(* IEC 61131-3 sources: sis-interlock-demo/tests/POUs/Generated/FB_CemGen01_Test, 41 files *)

(* ---- FB_CemGen01_Test.decl.st ---- *)
// AUTO-GENERATED by cemgen 1.0.0 — не редактировать: правьте матрицу и запустите
//   python -m cemgen generate <файл матрицы .csv или .xlsx>
// Матрица: SIS-V101-CEM, объект V-101, ревизия B от 2026-10-19, SHA-256 сетки df2ed4841a9453ca
// Назначение: набор coUnit: сценарии по матрице SIS-V101-CEM, тесты 1–40 (DESIGN.md, 12.4).
//             Ожидаемые значения — эталонная модель cemgen. Стенд FB_SisHarness — по экземпляру на
//             тест.
// Автор:      kr0nsch; код — генератор cemgen
// Версия:     1.0.0
// Документ:   docs/DESIGN.md, раздел «10. Генератор cemgen»; docs/cause_effect_matrix.md
// ВНИМАНИЕ:   код демонстрационный и не предназначен для систем безопасности. Реальная ПАЗ требует
//             определения SIL, сертифицированных аппаратных и программных средств и валидации по
//             ГОСТ Р МЭК 61511.
FUNCTION_BLOCK FB_CemGen01_Test EXTENDS coUnit.FB_TestSuite
VAR
    fbH001 : FB_SisHarness;   // Matrix_PSHH101Demand_TripsOwnEffects
    fbH002 : FB_SisHarness;   // Matrix_PSHH101Delay_TripsExactlyAtDelay
    fbH003 : FB_SisHarness;   // Matrix_PSHH101Override_Denied
    fbH004 : FB_SisHarness;   // Matrix_PSHH101Reset_OnlyAfterClear
    fbH005 : FB_SisHarness;   // Matrix_PSHH101ChannelInvalid_MatchesPolicy
    fbH006 : FB_SisHarness;   // Matrix_PSHH101Bypass_ExpiresBackToVoting
    fbH007 : FB_SisHarness;   // Matrix_PSLL101Demand_TripsOwnEffects
    fbH008 : FB_SisHarness;   // Matrix_PSLL101Delay_TripsExactlyAtDelay
    fbH009 : FB_SisHarness;   // Matrix_PSLL101Override_ExpiresThenTrips
    fbH010 : FB_SisHarness;   // Matrix_PSLL101Override_ClearsAfterConfirm
    fbH011 : FB_SisHarness;   // Matrix_PSLL101Override_DemandBackRestartsConfirm
    fbH012 : FB_SisHarness;   // Matrix_PSLL101Override_ExpiryBoundsConfirm
    fbH013 : FB_SisHarness;   // Matrix_PSLL101Override_ClearedThenDelayTrips
    fbH014 : FB_SisHarness;   // Matrix_PSLL101Reset_OnlyAfterClear
    fbH015 : FB_SisHarness;   // Matrix_PSLL101ChannelInvalid_MatchesPolicy
    fbH016 : FB_SisHarness;   // Matrix_PSLL101Bypass_ExpiresBackToVoting
    fbH017 : FB_SisHarness;   // Matrix_LSHH102Demand_TripsOwnEffects
    fbH018 : FB_SisHarness;   // Matrix_LSHH102Delay_TripsExactlyAtDelay
    fbH019 : FB_SisHarness;   // Matrix_LSHH102Override_Denied
    fbH020 : FB_SisHarness;   // Matrix_LSHH102Reset_OnlyAfterClear
    fbH021 : FB_SisHarness;   // Matrix_LSHH102ChannelInvalid_MatchesPolicy
    fbH022 : FB_SisHarness;   // Matrix_LSHH102Bypass_ExpiresBackToVoting
    fbH023 : FB_SisHarness;   // Matrix_LSLL102Demand_TripsOwnEffects
    fbH024 : FB_SisHarness;   // Matrix_LSLL102Delay_TripsExactlyAtDelay
    fbH025 : FB_SisHarness;   // Matrix_LSLL102Override_ExpiresThenTrips
    fbH026 : FB_SisHarness;   // Matrix_LSLL102Override_ClearsAfterConfirm
    fbH027 : FB_SisHarness;   // Matrix_LSLL102Override_DemandBackRestartsConfirm
    fbH028 : FB_SisHarness;   // Matrix_LSLL102Override_ExpiryBoundsConfirm
    fbH029 : FB_SisHarness;   // Matrix_LSLL102Override_ClearedThenDelayTrips
    fbH030 : FB_SisHarness;   // Matrix_LSLL102Reset_OnlyAfterClear
    fbH031 : FB_SisHarness;   // Matrix_LSLL102ChannelInvalid_MatchesPolicy
    fbH032 : FB_SisHarness;   // Matrix_LSLL102Bypass_ExpiresBackToVoting
    fbH033 : FB_SisHarness;   // Matrix_TSHH103Demand_TripsOwnEffects
    fbH034 : FB_SisHarness;   // Matrix_TSHH103Delay_TripsExactlyAtDelay
    fbH035 : FB_SisHarness;   // Matrix_TSHH103Override_Denied
    fbH036 : FB_SisHarness;   // Matrix_TSHH103Reset_OnlyAfterClear
    fbH037 : FB_SisHarness;   // Matrix_TSHH103ChannelInvalid_MatchesPolicy
    fbH038 : FB_SisHarness;   // Matrix_TSHH103Bypass_ExpiresBackToVoting
    fbH039 : FB_SisHarness;   // Matrix_ASHH104Demand_TripsOwnEffects
    fbH040 : FB_SisHarness;   // Matrix_ASHH104Delay_TripsExactlyAtDelay
END_VAR

(* ---- ASHH104DelayTripsExactlyAtDelay.method.decl.st ---- *)
// AUTO-GENERATED by cemgen 1.0.0 — не редактировать: правьте матрицу и запустите
//   python -m cemgen generate <файл матрицы .csv или .xlsx>
// Матрица: SIS-V101-CEM, объект V-101, ревизия B от 2026-10-19, SHA-256 сетки df2ed4841a9453ca
// Назначение: тест Matrix_ASHH104Delay_TripsExactlyAtDelay набора FB_CemGen01_Test (сценарий по
//             матрице, DESIGN.md, 12.4).
// Автор:      kr0nsch; код — генератор cemgen
// Версия:     1.0.0
// Документ:   docs/DESIGN.md, раздел «10. Генератор cemgen»; docs/cause_effect_matrix.md
// ВНИМАНИЕ:   код демонстрационный и не предназначен для систем безопасности. Реальная ПАЗ требует
//             определения SIL, сертифицированных аппаратных и программных средств и валидации по
//             ГОСТ Р МЭК 61511.
// Причина 6 ASHH104: требование в t0; на t0 + 2 с − шаг не зафиксирована, следствия под напряжением;
// ровно на t0 + 2 с — зафиксирована, ltFirstOut = t0 + задержка.
METHOD PRIVATE ASHH104DelayTripsExactlyAtDelay
VAR
    xArmed : BOOL;    // стенд взведён: все следствия под напряжением после сброса
    ltT0   : LTIME;   // момент t0 по подменному времени стенда
END_VAR

(* ---- ASHH104DemandTripsOwnEffects.method.decl.st ---- *)
// AUTO-GENERATED by cemgen 1.0.0 — не редактировать: правьте матрицу и запустите
//   python -m cemgen generate <файл матрицы .csv или .xlsx>
// Матрица: SIS-V101-CEM, объект V-101, ревизия B от 2026-10-19, SHA-256 сетки df2ed4841a9453ca
// Назначение: тест Matrix_ASHH104Demand_TripsOwnEffects набора FB_CemGen01_Test (сценарий по
//             матрице, DESIGN.md, 12.4).
// Автор:      kr0nsch; код — генератор cemgen
// Версия:     1.0.0
// Документ:   docs/DESIGN.md, раздел «10. Генератор cemgen»; docs/cause_effect_matrix.md
// ВНИМАНИЕ:   код демонстрационный и не предназначен для систем безопасности. Реальная ПАЗ требует
//             определения SIL, сертифицированных аппаратных и программных средств и валидации по
//             ГОСТ Р МЭК 61511.
// Причина 6 ASHH104 (2oo3, задержка 2 с): требование AT104A, AT104B, AT104C = 12,80 мА (55 % НКПР;
// уставка ≥ 50 % НКПР) отключает ESDV101, ESDV102, P101A, P101B, H101, UA110; остальные следствия под
// напряжением; первопричина ASHH104.
METHOD PRIVATE ASHH104DemandTripsOwnEffects
VAR
    xArmed : BOOL;   // стенд взведён: все следствия под напряжением после сброса
END_VAR

(* ---- LSHH102BypassExpiresBackToVoting.method.decl.st ---- *)
// AUTO-GENERATED by cemgen 1.0.0 — не редактировать: правьте матрицу и запустите
//   python -m cemgen generate <файл матрицы .csv или .xlsx>
// Матрица: SIS-V101-CEM, объект V-101, ревизия B от 2026-10-19, SHA-256 сетки df2ed4841a9453ca
// Назначение: тест Matrix_LSHH102Bypass_ExpiresBackToVoting набора FB_CemGen01_Test (сценарий по
//             матрице, DESIGN.md, 12.4).
// Автор:      kr0nsch; код — генератор cemgen
// Версия:     1.0.0
// Документ:   docs/DESIGN.md, раздел «10. Генератор cemgen»; docs/cause_effect_matrix.md
// ВНИМАНИЕ:   код демонстрационный и не предназначен для систем безопасности. Реальная ПАЗ требует
//             определения SIL, сертифицированных аппаратных и программных средств и валидации по
//             ГОСТ Р МЭК 61511.
// Причина 3 LSHH102: ключ разрешения байпасов, байпас LT102A → Active; канал недостоверен → Bypassed,
// не сработало; на t0 + 8 ч − шаг — Active; ровно на t0 + 8 ч — Expired, BypassExpired, канал Invalid;
// далее — по эталонной модели.
METHOD PRIVATE LSHH102BypassExpiresBackToVoting
VAR
    xArmed : BOOL;           // стенд взведён: все следствия под напряжением после сброса
    stVs   : ST_VotingSts;   // копия состояния группы голосования
END_VAR

(* ---- LSHH102ChannelInvalidMatchesPolicy.method.decl.st ---- *)
// AUTO-GENERATED by cemgen 1.0.0 — не редактировать: правьте матрицу и запустите
//   python -m cemgen generate <файл матрицы .csv или .xlsx>
// Матрица: SIS-V101-CEM, объект V-101, ревизия B от 2026-10-19, SHA-256 сетки df2ed4841a9453ca
// Назначение: тест Matrix_LSHH102ChannelInvalid_MatchesPolicy набора FB_CemGen01_Test (сценарий по
//             матрице, DESIGN.md, 12.4).
// Автор:      kr0nsch; код — генератор cemgen
// Версия:     1.0.0
// Документ:   docs/DESIGN.md, раздел «10. Генератор cemgen»; docs/cause_effect_matrix.md
// ВНИМАНИЕ:   код демонстрационный и не предназначен для систем безопасности. Реальная ПАЗ требует
//             определения SIL, сертифицированных аппаратных и программных средств и валидации по
//             ГОСТ Р МЭК 61511.
// Причина 3 LSHH102 (2oo3, DegradeAvailable): канал LT102A недостоверен → действующая схема и
// срабатывание по политике деградации; если не сработало — требование на LT102B → по эталонной модели.
METHOD PRIVATE LSHH102ChannelInvalidMatchesPolicy
VAR
    xArmed : BOOL;           // стенд взведён: все следствия под напряжением после сброса
    stVs   : ST_VotingSts;   // копия состояния группы голосования
END_VAR

(* ---- LSHH102DelayTripsExactlyAtDelay.method.decl.st ---- *)
// AUTO-GENERATED by cemgen 1.0.0 — не редактировать: правьте матрицу и запустите
//   python -m cemgen generate <файл матрицы .csv или .xlsx>
// Матрица: SIS-V101-CEM, объект V-101, ревизия B от 2026-10-19, SHA-256 сетки df2ed4841a9453ca
// Назначение: тест Matrix_LSHH102Delay_TripsExactlyAtDelay набора FB_CemGen01_Test (сценарий по
//             матрице, DESIGN.md, 12.4).
// Автор:      kr0nsch; код — генератор cemgen
// Версия:     1.0.0
// Документ:   docs/DESIGN.md, раздел «10. Генератор cemgen»; docs/cause_effect_matrix.md
// ВНИМАНИЕ:   код демонстрационный и не предназначен для систем безопасности. Реальная ПАЗ требует
//             определения SIL, сертифицированных аппаратных и программных средств и валидации по
//             ГОСТ Р МЭК 61511.
// Причина 3 LSHH102: требование в t0; на t0 + 3 с − шаг не зафиксирована, следствия под напряжением;
// ровно на t0 + 3 с — зафиксирована, ltFirstOut = t0 + задержка.
METHOD PRIVATE LSHH102DelayTripsExactlyAtDelay
VAR
    xArmed : BOOL;    // стенд взведён: все следствия под напряжением после сброса
    ltT0   : LTIME;   // момент t0 по подменному времени стенда
END_VAR

(* ---- LSHH102DemandTripsOwnEffects.method.decl.st ---- *)
// AUTO-GENERATED by cemgen 1.0.0 — не редактировать: правьте матрицу и запустите
//   python -m cemgen generate <файл матрицы .csv или .xlsx>
// Матрица: SIS-V101-CEM, объект V-101, ревизия B от 2026-10-19, SHA-256 сетки df2ed4841a9453ca
// Назначение: тест Matrix_LSHH102Demand_TripsOwnEffects набора FB_CemGen01_Test (сценарий по
//             матрице, DESIGN.md, 12.4).
// Автор:      kr0nsch; код — генератор cemgen
// Версия:     1.0.0
// Документ:   docs/DESIGN.md, раздел «10. Генератор cemgen»; docs/cause_effect_matrix.md
// ВНИМАНИЕ:   код демонстрационный и не предназначен для систем безопасности. Реальная ПАЗ требует
//             определения SIL, сертифицированных аппаратных и программных средств и валидации по
//             ГОСТ Р МЭК 61511.
// Причина 3 LSHH102 (2oo3, задержка 3 с): требование LT102A, LT102B, LT102C = 16,16 мА (1,824 м;
// уставка ≥ 1,8 м) отключает ESDV101, H101, UA110; остальные следствия под напряжением; первопричина
// LSHH102.
METHOD PRIVATE LSHH102DemandTripsOwnEffects
VAR
    xArmed : BOOL;   // стенд взведён: все следствия под напряжением после сброса
END_VAR

(* ---- LSHH102OverrideDenied.method.decl.st ---- *)
// AUTO-GENERATED by cemgen 1.0.0 — не редактировать: правьте матрицу и запустите
//   python -m cemgen generate <файл матрицы .csv или .xlsx>
// Матрица: SIS-V101-CEM, объект V-101, ревизия B от 2026-10-19, SHA-256 сетки df2ed4841a9453ca
// Назначение: тест Matrix_LSHH102Override_Denied набора FB_CemGen01_Test (сценарий по матрице,
//             DESIGN.md, 12.4).
// Автор:      kr0nsch; код — генератор cemgen
// Версия:     1.0.0
// Документ:   docs/DESIGN.md, раздел «10. Генератор cemgen»; docs/cause_effect_matrix.md
// ВНИМАНИЕ:   код демонстрационный и не предназначен для систем безопасности. Реальная ПАЗ требует
//             определения SIL, сертифицированных аппаратных и программных средств и валидации по
//             ГОСТ Р МЭК 61511.
// Причина 3 LSHH102 без разрешённого обхода: ключ разрешения обходов, запрос → последнее событие
// OverrideDenied, обхода нет; требование → срабатывание после задержки.
METHOD PRIVATE LSHH102OverrideDenied
VAR
    xArmed : BOOL;          // стенд взведён: все следствия под напряжением после сброса
    stEv   : ST_SisEvent;   // последнее событие журнала
END_VAR

(* ---- LSHH102ResetOnlyAfterClear.method.decl.st ---- *)
// AUTO-GENERATED by cemgen 1.0.0 — не редактировать: правьте матрицу и запустите
//   python -m cemgen generate <файл матрицы .csv или .xlsx>
// Матрица: SIS-V101-CEM, объект V-101, ревизия B от 2026-10-19, SHA-256 сетки df2ed4841a9453ca
// Назначение: тест Matrix_LSHH102Reset_OnlyAfterClear набора FB_CemGen01_Test (сценарий по матрице,
//             DESIGN.md, 12.4).
// Автор:      kr0nsch; код — генератор cemgen
// Версия:     1.0.0
// Документ:   docs/DESIGN.md, раздел «10. Генератор cemgen»; docs/cause_effect_matrix.md
// ВНИМАНИЕ:   код демонстрационный и не предназначен для систем безопасности. Реальная ПАЗ требует
//             определения SIL, сертифицированных аппаратных и программных средств и валидации по
//             ГОСТ Р МЭК 61511.
// Причина 3 LSHH102: срабатывание; сброс при требовании → ResetDenied, блокирует LSHH102, следствия
// обесточены; норма → следствия всё ещё обесточены (фиксация); сброс → все следствия под напряжением.
METHOD PRIVATE LSHH102ResetOnlyAfterClear
VAR
    xArmed : BOOL;          // стенд взведён: все следствия под напряжением после сброса
    stEv   : ST_SisEvent;   // последнее событие журнала
END_VAR

(* ---- LSLL102BypassExpiresBackToVoting.method.decl.st ---- *)
// AUTO-GENERATED by cemgen 1.0.0 — не редактировать: правьте матрицу и запустите
//   python -m cemgen generate <файл матрицы .csv или .xlsx>
// Матрица: SIS-V101-CEM, объект V-101, ревизия B от 2026-10-19, SHA-256 сетки df2ed4841a9453ca
// Назначение: тест Matrix_LSLL102Bypass_ExpiresBackToVoting набора FB_CemGen01_Test (сценарий по
//             матрице, DESIGN.md, 12.4).
// Автор:      kr0nsch; код — генератор cemgen
// Версия:     1.0.0
// Документ:   docs/DESIGN.md, раздел «10. Генератор cemgen»; docs/cause_effect_matrix.md
// ВНИМАНИЕ:   код демонстрационный и не предназначен для систем безопасности. Реальная ПАЗ требует
//             определения SIL, сертифицированных аппаратных и программных средств и валидации по
//             ГОСТ Р МЭК 61511.
// Причина 4 LSLL102: ключ разрешения байпасов, байпас LT102A → Active; канал недостоверен → Bypassed,
// не сработало; на t0 + 8 ч − шаг — Active; ровно на t0 + 8 ч — Expired, BypassExpired, канал Invalid;
// далее — по эталонной модели.
METHOD PRIVATE LSLL102BypassExpiresBackToVoting
VAR
    xArmed : BOOL;           // стенд взведён: все следствия под напряжением после сброса
    stVs   : ST_VotingSts;   // копия состояния группы голосования
END_VAR

(* ---- LSLL102ChannelInvalidMatchesPolicy.method.decl.st ---- *)
// AUTO-GENERATED by cemgen 1.0.0 — не редактировать: правьте матрицу и запустите
//   python -m cemgen generate <файл матрицы .csv или .xlsx>
// Матрица: SIS-V101-CEM, объект V-101, ревизия B от 2026-10-19, SHA-256 сетки df2ed4841a9453ca
// Назначение: тест Matrix_LSLL102ChannelInvalid_MatchesPolicy набора FB_CemGen01_Test (сценарий по
//             матрице, DESIGN.md, 12.4).
// Автор:      kr0nsch; код — генератор cemgen
// Версия:     1.0.0
// Документ:   docs/DESIGN.md, раздел «10. Генератор cemgen»; docs/cause_effect_matrix.md
// ВНИМАНИЕ:   код демонстрационный и не предназначен для систем безопасности. Реальная ПАЗ требует
//             определения SIL, сертифицированных аппаратных и программных средств и валидации по
//             ГОСТ Р МЭК 61511.
// Причина 4 LSLL102 (2oo3, DegradeAvailable): канал LT102A недостоверен → действующая схема и
// срабатывание по политике деградации; если не сработало — требование на LT102B → по эталонной модели.
METHOD PRIVATE LSLL102ChannelInvalidMatchesPolicy
VAR
    xArmed : BOOL;           // стенд взведён: все следствия под напряжением после сброса
    stVs   : ST_VotingSts;   // копия состояния группы голосования
END_VAR

(* ---- LSLL102DelayTripsExactlyAtDelay.method.decl.st ---- *)
// AUTO-GENERATED by cemgen 1.0.0 — не редактировать: правьте матрицу и запустите
//   python -m cemgen generate <файл матрицы .csv или .xlsx>
// Матрица: SIS-V101-CEM, объект V-101, ревизия B от 2026-10-19, SHA-256 сетки df2ed4841a9453ca
// Назначение: тест Matrix_LSLL102Delay_TripsExactlyAtDelay набора FB_CemGen01_Test (сценарий по
//             матрице, DESIGN.md, 12.4).
// Автор:      kr0nsch; код — генератор cemgen
// Версия:     1.0.0
// Документ:   docs/DESIGN.md, раздел «10. Генератор cemgen»; docs/cause_effect_matrix.md
// ВНИМАНИЕ:   код демонстрационный и не предназначен для систем безопасности. Реальная ПАЗ требует
//             определения SIL, сертифицированных аппаратных и программных средств и валидации по
//             ГОСТ Р МЭК 61511.
// Причина 4 LSLL102: требование в t0; на t0 + 5 с − шаг не зафиксирована, следствия под напряжением;
// ровно на t0 + 5 с — зафиксирована, ltFirstOut = t0 + задержка.
METHOD PRIVATE LSLL102DelayTripsExactlyAtDelay
VAR
    xArmed : BOOL;    // стенд взведён: все следствия под напряжением после сброса
    ltT0   : LTIME;   // момент t0 по подменному времени стенда
END_VAR

(* ---- LSLL102DemandTripsOwnEffects.method.decl.st ---- *)
// AUTO-GENERATED by cemgen 1.0.0 — не редактировать: правьте матрицу и запустите
//   python -m cemgen generate <файл матрицы .csv или .xlsx>
// Матрица: SIS-V101-CEM, объект V-101, ревизия B от 2026-10-19, SHA-256 сетки df2ed4841a9453ca
// Назначение: тест Matrix_LSLL102Demand_TripsOwnEffects набора FB_CemGen01_Test (сценарий по
//             матрице, DESIGN.md, 12.4).
// Автор:      kr0nsch; код — генератор cemgen
// Версия:     1.0.0
// Документ:   docs/DESIGN.md, раздел «10. Генератор cemgen»; docs/cause_effect_matrix.md
// ВНИМАНИЕ:   код демонстрационный и не предназначен для систем безопасности. Реальная ПАЗ требует
//             определения SIL, сертифицированных аппаратных и программных средств и валидации по
//             ГОСТ Р МЭК 61511.
// Причина 4 LSLL102 (2oo3, задержка 5 с): требование LT102A, LT102B, LT102C = 7,17 мА (0,476 м;
// уставка ≤ 0,5 м) отключает ESDV102, P101A, P101B, H101, UA110; остальные следствия под напряжением;
// первопричина LSLL102.
METHOD PRIVATE LSLL102DemandTripsOwnEffects
VAR
    xArmed : BOOL;   // стенд взведён: все следствия под напряжением после сброса
END_VAR

(* ---- LSLL102OverrideClearedThenDelayTrips.method.decl.st ---- *)
// AUTO-GENERATED by cemgen 1.0.0 — не редактировать: правьте матрицу и запустите
//   python -m cemgen generate <файл матрицы .csv или .xlsx>
// Матрица: SIS-V101-CEM, объект V-101, ревизия B от 2026-10-19, SHA-256 сетки df2ed4841a9453ca
// Назначение: тест Matrix_LSLL102Override_ClearedThenDelayTrips набора FB_CemGen01_Test (сценарий
//             по матрице, DESIGN.md, 12.4).
// Автор:      kr0nsch; код — генератор cemgen
// Версия:     1.0.0
// Документ:   docs/DESIGN.md, раздел «10. Генератор cemgen»; docs/cause_effect_matrix.md
// ВНИМАНИЕ:   код демонстрационный и не предназначен для систем безопасности. Реальная ПАЗ требует
//             определения SIL, сертифицированных аппаратных и программных средств и валидации по
//             ГОСТ Р МЭК 61511.
// Причина 4 LSLL102 с задержкой 5 с: пусковой обход и требование в t0; через 5 с причина активна под
// обходом, не зафиксирована; норма; через 1 мин — OverrideCleared; требование в t2 — на t2 + 5 с − шаг
// не зафиксирована (задержка отсчитывается заново), на t2 + 5 с — зафиксирована, первопричина LSLL102.
METHOD PRIVATE LSLL102OverrideClearedThenDelayTrips
VAR
    xArmed : BOOL;    // стенд взведён: все следствия под напряжением после сброса
    ltT0   : LTIME;   // момент t2 по подменному времени стенда
END_VAR

(* ---- LSLL102OverrideClearsAfterConfirm.method.decl.st ---- *)
// AUTO-GENERATED by cemgen 1.0.0 — не редактировать: правьте матрицу и запустите
//   python -m cemgen generate <файл матрицы .csv или .xlsx>
// Матрица: SIS-V101-CEM, объект V-101, ревизия B от 2026-10-19, SHA-256 сетки df2ed4841a9453ca
// Назначение: тест Matrix_LSLL102Override_ClearsAfterConfirm набора FB_CemGen01_Test (сценарий по
//             матрице, DESIGN.md, 12.4).
// Автор:      kr0nsch; код — генератор cemgen
// Версия:     1.0.0
// Документ:   docs/DESIGN.md, раздел «10. Генератор cemgen»; docs/cause_effect_matrix.md
// ВНИМАНИЕ:   код демонстрационный и не предназначен для систем безопасности. Реальная ПАЗ требует
//             определения SIL, сертифицированных аппаратных и программных средств и валидации по
//             ГОСТ Р МЭК 61511.
// Причина 4 LSLL102: пусковой обход и требование в t0; норма с t1 = t0 + шаг; на t1 + 1 мин − шаг
// обход действует; ровно на t1 + 1 мин (подтверждение нормы) — OverrideCleared, обхода нет, причина не
// зафиксирована, следствия под напряжением (R-12).
METHOD PRIVATE LSLL102OverrideClearsAfterConfirm
VAR
    xArmed : BOOL;   // стенд взведён: все следствия под напряжением после сброса
END_VAR

(* ---- LSLL102OverrideDemandBackRestartsConfirm.method.decl.st ---- *)
// AUTO-GENERATED by cemgen 1.0.0 — не редактировать: правьте матрицу и запустите
//   python -m cemgen generate <файл матрицы .csv или .xlsx>
// Матрица: SIS-V101-CEM, объект V-101, ревизия B от 2026-10-19, SHA-256 сетки df2ed4841a9453ca
// Назначение: тест Matrix_LSLL102Override_DemandBackRestartsConfirm набора FB_CemGen01_Test
//             (сценарий по матрице, DESIGN.md, 12.4).
// Автор:      kr0nsch; код — генератор cemgen
// Версия:     1.0.0
// Документ:   docs/DESIGN.md, раздел «10. Генератор cemgen»; docs/cause_effect_matrix.md
// ВНИМАНИЕ:   код демонстрационный и не предназначен для систем безопасности. Реальная ПАЗ требует
//             определения SIL, сертифицированных аппаратных и программных средств и валидации по
//             ГОСТ Р МЭК 61511.
// Причина 4 LSLL102: пусковой обход и требование в t0; норма с t1; ровно на t1 + 1 мин, когда обход
// снялся бы, требование снова — обход действует, подтверждение нормы сброшено; норма с t2; на t2 + 1
// мин − шаг обход действует; на t2 + 1 мин — OverrideCleared.
METHOD PRIVATE LSLL102OverrideDemandBackRestartsConfirm
VAR
    xArmed : BOOL;   // стенд взведён: все следствия под напряжением после сброса
END_VAR

(* ---- LSLL102OverrideExpiresThenTrips.method.decl.st ---- *)
// AUTO-GENERATED by cemgen 1.0.0 — не редактировать: правьте матрицу и запустите
//   python -m cemgen generate <файл матрицы .csv или .xlsx>
// Матрица: SIS-V101-CEM, объект V-101, ревизия B от 2026-10-19, SHA-256 сетки df2ed4841a9453ca
// Назначение: тест Matrix_LSLL102Override_ExpiresThenTrips набора FB_CemGen01_Test (сценарий по
//             матрице, DESIGN.md, 12.4).
// Автор:      kr0nsch; код — генератор cemgen
// Версия:     1.0.0
// Документ:   docs/DESIGN.md, раздел «10. Генератор cemgen»; docs/cause_effect_matrix.md
// ВНИМАНИЕ:   код демонстрационный и не предназначен для систем безопасности. Реальная ПАЗ требует
//             определения SIL, сертифицированных аппаратных и программных средств и валидации по
//             ГОСТ Р МЭК 61511.
// Причина 4 LSLL102: ключ разрешения обходов, запрос пускового обхода и требование в одном вызове t0;
// до t0 + 30 мин − шаг обход действует, причина не зафиксирована; ровно на t0 + 30 мин —
// OverrideExpired, фиксация, первопричина LSLL102.
METHOD PRIVATE LSLL102OverrideExpiresThenTrips
VAR
    xArmed : BOOL;   // стенд взведён: все следствия под напряжением после сброса
END_VAR

(* ---- LSLL102OverrideExpiryBoundsConfirm.method.decl.st ---- *)
// AUTO-GENERATED by cemgen 1.0.0 — не редактировать: правьте матрицу и запустите
//   python -m cemgen generate <файл матрицы .csv или .xlsx>
// Матрица: SIS-V101-CEM, объект V-101, ревизия B от 2026-10-19, SHA-256 сетки df2ed4841a9453ca
// Назначение: тест Matrix_LSLL102Override_ExpiryBoundsConfirm набора FB_CemGen01_Test (сценарий по
//             матрице, DESIGN.md, 12.4).
// Автор:      kr0nsch; код — генератор cemgen
// Версия:     1.0.0
// Документ:   docs/DESIGN.md, раздел «10. Генератор cemgen»; docs/cause_effect_matrix.md
// ВНИМАНИЕ:   код демонстрационный и не предназначен для систем безопасности. Реальная ПАЗ требует
//             определения SIL, сертифицированных аппаратных и программных средств и валидации по
//             ГОСТ Р МЭК 61511.
// Причина 4 LSLL102: пусковой обход и требование в t0; норма с t0 + 29 мин + шаг — подтверждение (1
// мин) закончилось бы после срока; на t0 + 30 мин − шаг обход действует; ровно на t0 + 30 мин —
// OverrideExpired (срок — верхняя граница), OverrideCleared нет, причина не зафиксирована (требования
// нет).
METHOD PRIVATE LSLL102OverrideExpiryBoundsConfirm
VAR
    xArmed : BOOL;   // стенд взведён: все следствия под напряжением после сброса
END_VAR

(* ---- LSLL102ResetOnlyAfterClear.method.decl.st ---- *)
// AUTO-GENERATED by cemgen 1.0.0 — не редактировать: правьте матрицу и запустите
//   python -m cemgen generate <файл матрицы .csv или .xlsx>
// Матрица: SIS-V101-CEM, объект V-101, ревизия B от 2026-10-19, SHA-256 сетки df2ed4841a9453ca
// Назначение: тест Matrix_LSLL102Reset_OnlyAfterClear набора FB_CemGen01_Test (сценарий по матрице,
//             DESIGN.md, 12.4).
// Автор:      kr0nsch; код — генератор cemgen
// Версия:     1.0.0
// Документ:   docs/DESIGN.md, раздел «10. Генератор cemgen»; docs/cause_effect_matrix.md
// ВНИМАНИЕ:   код демонстрационный и не предназначен для систем безопасности. Реальная ПАЗ требует
//             определения SIL, сертифицированных аппаратных и программных средств и валидации по
//             ГОСТ Р МЭК 61511.
// Причина 4 LSLL102: срабатывание; сброс при требовании → ResetDenied, блокирует LSLL102, следствия
// обесточены; норма → следствия всё ещё обесточены (фиксация); сброс → все следствия под напряжением.
METHOD PRIVATE LSLL102ResetOnlyAfterClear
VAR
    xArmed : BOOL;          // стенд взведён: все следствия под напряжением после сброса
    stEv   : ST_SisEvent;   // последнее событие журнала
END_VAR

(* ---- PSHH101BypassExpiresBackToVoting.method.decl.st ---- *)
// AUTO-GENERATED by cemgen 1.0.0 — не редактировать: правьте матрицу и запустите
//   python -m cemgen generate <файл матрицы .csv или .xlsx>
// Матрица: SIS-V101-CEM, объект V-101, ревизия B от 2026-10-19, SHA-256 сетки df2ed4841a9453ca
// Назначение: тест Matrix_PSHH101Bypass_ExpiresBackToVoting набора FB_CemGen01_Test (сценарий по
//             матрице, DESIGN.md, 12.4).
// Автор:      kr0nsch; код — генератор cemgen
// Версия:     1.0.0
// Документ:   docs/DESIGN.md, раздел «10. Генератор cemgen»; docs/cause_effect_matrix.md
// ВНИМАНИЕ:   код демонстрационный и не предназначен для систем безопасности. Реальная ПАЗ требует
//             определения SIL, сертифицированных аппаратных и программных средств и валидации по
//             ГОСТ Р МЭК 61511.
// Причина 1 PSHH101: ключ разрешения байпасов, байпас PT101A → Active; канал недостоверен → Bypassed,
// не сработало; на t0 + 8 ч − шаг — Active; ровно на t0 + 8 ч — Expired, BypassExpired, канал Invalid;
// далее — по эталонной модели.
METHOD PRIVATE PSHH101BypassExpiresBackToVoting
VAR
    xArmed : BOOL;           // стенд взведён: все следствия под напряжением после сброса
    stVs   : ST_VotingSts;   // копия состояния группы голосования
END_VAR

(* ---- PSHH101ChannelInvalidMatchesPolicy.method.decl.st ---- *)
// AUTO-GENERATED by cemgen 1.0.0 — не редактировать: правьте матрицу и запустите
//   python -m cemgen generate <файл матрицы .csv или .xlsx>
// Матрица: SIS-V101-CEM, объект V-101, ревизия B от 2026-10-19, SHA-256 сетки df2ed4841a9453ca
// Назначение: тест Matrix_PSHH101ChannelInvalid_MatchesPolicy набора FB_CemGen01_Test (сценарий по
//             матрице, DESIGN.md, 12.4).
// Автор:      kr0nsch; код — генератор cemgen
// Версия:     1.0.0
// Документ:   docs/DESIGN.md, раздел «10. Генератор cemgen»; docs/cause_effect_matrix.md
// ВНИМАНИЕ:   код демонстрационный и не предназначен для систем безопасности. Реальная ПАЗ требует
//             определения SIL, сертифицированных аппаратных и программных средств и валидации по
//             ГОСТ Р МЭК 61511.
// Причина 1 PSHH101 (2oo3, VoteTrip): канал PT101A недостоверен → действующая схема и срабатывание по
// политике деградации; если не сработало — требование на PT101B → по эталонной модели.
METHOD PRIVATE PSHH101ChannelInvalidMatchesPolicy
VAR
    xArmed : BOOL;           // стенд взведён: все следствия под напряжением после сброса
    stVs   : ST_VotingSts;   // копия состояния группы голосования
END_VAR

(* ---- PSHH101DelayTripsExactlyAtDelay.method.decl.st ---- *)
// AUTO-GENERATED by cemgen 1.0.0 — не редактировать: правьте матрицу и запустите
//   python -m cemgen generate <файл матрицы .csv или .xlsx>
// Матрица: SIS-V101-CEM, объект V-101, ревизия B от 2026-10-19, SHA-256 сетки df2ed4841a9453ca
// Назначение: тест Matrix_PSHH101Delay_TripsExactlyAtDelay набора FB_CemGen01_Test (сценарий по
//             матрице, DESIGN.md, 12.4).
// Автор:      kr0nsch; код — генератор cemgen
// Версия:     1.0.0
// Документ:   docs/DESIGN.md, раздел «10. Генератор cemgen»; docs/cause_effect_matrix.md
// ВНИМАНИЕ:   код демонстрационный и не предназначен для систем безопасности. Реальная ПАЗ требует
//             определения SIL, сертифицированных аппаратных и программных средств и валидации по
//             ГОСТ Р МЭК 61511.
// Причина 1 PSHH101: требование в t0; на t0 + 2 с − шаг не зафиксирована, следствия под напряжением;
// ровно на t0 + 2 с — зафиксирована, ltFirstOut = t0 + задержка.
METHOD PRIVATE PSHH101DelayTripsExactlyAtDelay
VAR
    xArmed : BOOL;    // стенд взведён: все следствия под напряжением после сброса
    ltT0   : LTIME;   // момент t0 по подменному времени стенда
END_VAR

(* ---- PSHH101DemandTripsOwnEffects.method.decl.st ---- *)
// AUTO-GENERATED by cemgen 1.0.0 — не редактировать: правьте матрицу и запустите
//   python -m cemgen generate <файл матрицы .csv или .xlsx>
// Матрица: SIS-V101-CEM, объект V-101, ревизия B от 2026-10-19, SHA-256 сетки df2ed4841a9453ca
// Назначение: тест Matrix_PSHH101Demand_TripsOwnEffects набора FB_CemGen01_Test (сценарий по
//             матрице, DESIGN.md, 12.4).
// Автор:      kr0nsch; код — генератор cemgen
// Версия:     1.0.0
// Документ:   docs/DESIGN.md, раздел «10. Генератор cemgen»; docs/cause_effect_matrix.md
// ВНИМАНИЕ:   код демонстрационный и не предназначен для систем безопасности. Реальная ПАЗ требует
//             определения SIL, сертифицированных аппаратных и программных средств и валидации по
//             ГОСТ Р МЭК 61511.
// Причина 1 PSHH101 (2oo3, задержка 2 с): требование PT101A, PT101B, PT101C = 13,20 мА (0,92 МПа;
// уставка ≥ 0,9 МПа) отключает ESDV101, H101, UA110; остальные следствия под напряжением; первопричина
// PSHH101.
METHOD PRIVATE PSHH101DemandTripsOwnEffects
VAR
    xArmed : BOOL;   // стенд взведён: все следствия под напряжением после сброса
END_VAR

(* ---- PSHH101OverrideDenied.method.decl.st ---- *)
// AUTO-GENERATED by cemgen 1.0.0 — не редактировать: правьте матрицу и запустите
//   python -m cemgen generate <файл матрицы .csv или .xlsx>
// Матрица: SIS-V101-CEM, объект V-101, ревизия B от 2026-10-19, SHA-256 сетки df2ed4841a9453ca
// Назначение: тест Matrix_PSHH101Override_Denied набора FB_CemGen01_Test (сценарий по матрице,
//             DESIGN.md, 12.4).
// Автор:      kr0nsch; код — генератор cemgen
// Версия:     1.0.0
// Документ:   docs/DESIGN.md, раздел «10. Генератор cemgen»; docs/cause_effect_matrix.md
// ВНИМАНИЕ:   код демонстрационный и не предназначен для систем безопасности. Реальная ПАЗ требует
//             определения SIL, сертифицированных аппаратных и программных средств и валидации по
//             ГОСТ Р МЭК 61511.
// Причина 1 PSHH101 без разрешённого обхода: ключ разрешения обходов, запрос → последнее событие
// OverrideDenied, обхода нет; требование → срабатывание после задержки.
METHOD PRIVATE PSHH101OverrideDenied
VAR
    xArmed : BOOL;          // стенд взведён: все следствия под напряжением после сброса
    stEv   : ST_SisEvent;   // последнее событие журнала
END_VAR

(* ---- PSHH101ResetOnlyAfterClear.method.decl.st ---- *)
// AUTO-GENERATED by cemgen 1.0.0 — не редактировать: правьте матрицу и запустите
//   python -m cemgen generate <файл матрицы .csv или .xlsx>
// Матрица: SIS-V101-CEM, объект V-101, ревизия B от 2026-10-19, SHA-256 сетки df2ed4841a9453ca
// Назначение: тест Matrix_PSHH101Reset_OnlyAfterClear набора FB_CemGen01_Test (сценарий по матрице,
//             DESIGN.md, 12.4).
// Автор:      kr0nsch; код — генератор cemgen
// Версия:     1.0.0
// Документ:   docs/DESIGN.md, раздел «10. Генератор cemgen»; docs/cause_effect_matrix.md
// ВНИМАНИЕ:   код демонстрационный и не предназначен для систем безопасности. Реальная ПАЗ требует
//             определения SIL, сертифицированных аппаратных и программных средств и валидации по
//             ГОСТ Р МЭК 61511.
// Причина 1 PSHH101: срабатывание; сброс при требовании → ResetDenied, блокирует PSHH101, следствия
// обесточены; норма → следствия всё ещё обесточены (фиксация); сброс → все следствия под напряжением.
METHOD PRIVATE PSHH101ResetOnlyAfterClear
VAR
    xArmed : BOOL;          // стенд взведён: все следствия под напряжением после сброса
    stEv   : ST_SisEvent;   // последнее событие журнала
END_VAR

(* ---- PSLL101BypassExpiresBackToVoting.method.decl.st ---- *)
// AUTO-GENERATED by cemgen 1.0.0 — не редактировать: правьте матрицу и запустите
//   python -m cemgen generate <файл матрицы .csv или .xlsx>
// Матрица: SIS-V101-CEM, объект V-101, ревизия B от 2026-10-19, SHA-256 сетки df2ed4841a9453ca
// Назначение: тест Matrix_PSLL101Bypass_ExpiresBackToVoting набора FB_CemGen01_Test (сценарий по
//             матрице, DESIGN.md, 12.4).
// Автор:      kr0nsch; код — генератор cemgen
// Версия:     1.0.0
// Документ:   docs/DESIGN.md, раздел «10. Генератор cemgen»; docs/cause_effect_matrix.md
// ВНИМАНИЕ:   код демонстрационный и не предназначен для систем безопасности. Реальная ПАЗ требует
//             определения SIL, сертифицированных аппаратных и программных средств и валидации по
//             ГОСТ Р МЭК 61511.
// Причина 2 PSLL101: ключ разрешения байпасов, байпас PT101A → Active; канал недостоверен → Bypassed,
// не сработало; на t0 + 8 ч − шаг — Active; ровно на t0 + 8 ч — Expired, BypassExpired, канал Invalid;
// далее — по эталонной модели.
METHOD PRIVATE PSLL101BypassExpiresBackToVoting
VAR
    xArmed : BOOL;           // стенд взведён: все следствия под напряжением после сброса
    stVs   : ST_VotingSts;   // копия состояния группы голосования
END_VAR

(* ---- PSLL101ChannelInvalidMatchesPolicy.method.decl.st ---- *)
// AUTO-GENERATED by cemgen 1.0.0 — не редактировать: правьте матрицу и запустите
//   python -m cemgen generate <файл матрицы .csv или .xlsx>
// Матрица: SIS-V101-CEM, объект V-101, ревизия B от 2026-10-19, SHA-256 сетки df2ed4841a9453ca
// Назначение: тест Matrix_PSLL101ChannelInvalid_MatchesPolicy набора FB_CemGen01_Test (сценарий по
//             матрице, DESIGN.md, 12.4).
// Автор:      kr0nsch; код — генератор cemgen
// Версия:     1.0.0
// Документ:   docs/DESIGN.md, раздел «10. Генератор cemgen»; docs/cause_effect_matrix.md
// ВНИМАНИЕ:   код демонстрационный и не предназначен для систем безопасности. Реальная ПАЗ требует
//             определения SIL, сертифицированных аппаратных и программных средств и валидации по
//             ГОСТ Р МЭК 61511.
// Причина 2 PSLL101 (2oo3, VoteTrip): канал PT101A недостоверен → действующая схема и срабатывание по
// политике деградации; если не сработало — требование на PT101B → по эталонной модели.
METHOD PRIVATE PSLL101ChannelInvalidMatchesPolicy
VAR
    xArmed : BOOL;           // стенд взведён: все следствия под напряжением после сброса
    stVs   : ST_VotingSts;   // копия состояния группы голосования
END_VAR

(* ---- PSLL101DelayTripsExactlyAtDelay.method.decl.st ---- *)
// AUTO-GENERATED by cemgen 1.0.0 — не редактировать: правьте матрицу и запустите
//   python -m cemgen generate <файл матрицы .csv или .xlsx>
// Матрица: SIS-V101-CEM, объект V-101, ревизия B от 2026-10-19, SHA-256 сетки df2ed4841a9453ca
// Назначение: тест Matrix_PSLL101Delay_TripsExactlyAtDelay набора FB_CemGen01_Test (сценарий по
//             матрице, DESIGN.md, 12.4).
// Автор:      kr0nsch; код — генератор cemgen
// Версия:     1.0.0
// Документ:   docs/DESIGN.md, раздел «10. Генератор cemgen»; docs/cause_effect_matrix.md
// ВНИМАНИЕ:   код демонстрационный и не предназначен для систем безопасности. Реальная ПАЗ требует
//             определения SIL, сертифицированных аппаратных и программных средств и валидации по
//             ГОСТ Р МЭК 61511.
// Причина 2 PSLL101: требование в t0; на t0 + 5 с − шаг не зафиксирована, следствия под напряжением;
// ровно на t0 + 5 с — зафиксирована, ltFirstOut = t0 + задержка.
METHOD PRIVATE PSLL101DelayTripsExactlyAtDelay
VAR
    xArmed : BOOL;    // стенд взведён: все следствия под напряжением после сброса
    ltT0   : LTIME;   // момент t0 по подменному времени стенда
END_VAR

(* ---- PSLL101DemandTripsOwnEffects.method.decl.st ---- *)
// AUTO-GENERATED by cemgen 1.0.0 — не редактировать: правьте матрицу и запустите
//   python -m cemgen generate <файл матрицы .csv или .xlsx>
// Матрица: SIS-V101-CEM, объект V-101, ревизия B от 2026-10-19, SHA-256 сетки df2ed4841a9453ca
// Назначение: тест Matrix_PSLL101Demand_TripsOwnEffects набора FB_CemGen01_Test (сценарий по
//             матрице, DESIGN.md, 12.4).
// Автор:      kr0nsch; код — генератор cemgen
// Версия:     1.0.0
// Документ:   docs/DESIGN.md, раздел «10. Генератор cemgen»; docs/cause_effect_matrix.md
// ВНИМАНИЕ:   код демонстрационный и не предназначен для систем безопасности. Реальная ПАЗ требует
//             определения SIL, сертифицированных аппаратных и программных средств и валидации по
//             ГОСТ Р МЭК 61511.
// Причина 2 PSLL101 (2oo3, задержка 5 с): требование PT101A, PT101B, PT101C = 5,30 мА (0,13 МПа;
// уставка ≤ 0,15 МПа) отключает ESDV101, ESDV102, P101A, P101B, H101, UA110; остальные следствия под
// напряжением; первопричина PSLL101.
METHOD PRIVATE PSLL101DemandTripsOwnEffects
VAR
    xArmed : BOOL;   // стенд взведён: все следствия под напряжением после сброса
END_VAR

(* ---- PSLL101OverrideClearedThenDelayTrips.method.decl.st ---- *)
// AUTO-GENERATED by cemgen 1.0.0 — не редактировать: правьте матрицу и запустите
//   python -m cemgen generate <файл матрицы .csv или .xlsx>
// Матрица: SIS-V101-CEM, объект V-101, ревизия B от 2026-10-19, SHA-256 сетки df2ed4841a9453ca
// Назначение: тест Matrix_PSLL101Override_ClearedThenDelayTrips набора FB_CemGen01_Test (сценарий
//             по матрице, DESIGN.md, 12.4).
// Автор:      kr0nsch; код — генератор cemgen
// Версия:     1.0.0
// Документ:   docs/DESIGN.md, раздел «10. Генератор cemgen»; docs/cause_effect_matrix.md
// ВНИМАНИЕ:   код демонстрационный и не предназначен для систем безопасности. Реальная ПАЗ требует
//             определения SIL, сертифицированных аппаратных и программных средств и валидации по
//             ГОСТ Р МЭК 61511.
// Причина 2 PSLL101 с задержкой 5 с: пусковой обход и требование в t0; через 5 с причина активна под
// обходом, не зафиксирована; норма; через 30 с — OverrideCleared; требование в t2 — на t2 + 5 с − шаг
// не зафиксирована (задержка отсчитывается заново), на t2 + 5 с — зафиксирована, первопричина PSLL101.
METHOD PRIVATE PSLL101OverrideClearedThenDelayTrips
VAR
    xArmed : BOOL;    // стенд взведён: все следствия под напряжением после сброса
    ltT0   : LTIME;   // момент t2 по подменному времени стенда
END_VAR

(* ---- PSLL101OverrideClearsAfterConfirm.method.decl.st ---- *)
// AUTO-GENERATED by cemgen 1.0.0 — не редактировать: правьте матрицу и запустите
//   python -m cemgen generate <файл матрицы .csv или .xlsx>
// Матрица: SIS-V101-CEM, объект V-101, ревизия B от 2026-10-19, SHA-256 сетки df2ed4841a9453ca
// Назначение: тест Matrix_PSLL101Override_ClearsAfterConfirm набора FB_CemGen01_Test (сценарий по
//             матрице, DESIGN.md, 12.4).
// Автор:      kr0nsch; код — генератор cemgen
// Версия:     1.0.0
// Документ:   docs/DESIGN.md, раздел «10. Генератор cemgen»; docs/cause_effect_matrix.md
// ВНИМАНИЕ:   код демонстрационный и не предназначен для систем безопасности. Реальная ПАЗ требует
//             определения SIL, сертифицированных аппаратных и программных средств и валидации по
//             ГОСТ Р МЭК 61511.
// Причина 2 PSLL101: пусковой обход и требование в t0; норма с t1 = t0 + шаг; на t1 + 30 с − шаг обход
// действует; ровно на t1 + 30 с (подтверждение нормы) — OverrideCleared, обхода нет, причина не
// зафиксирована, следствия под напряжением (R-12).
METHOD PRIVATE PSLL101OverrideClearsAfterConfirm
VAR
    xArmed : BOOL;   // стенд взведён: все следствия под напряжением после сброса
END_VAR

(* ---- PSLL101OverrideDemandBackRestartsConfirm.method.decl.st ---- *)
// AUTO-GENERATED by cemgen 1.0.0 — не редактировать: правьте матрицу и запустите
//   python -m cemgen generate <файл матрицы .csv или .xlsx>
// Матрица: SIS-V101-CEM, объект V-101, ревизия B от 2026-10-19, SHA-256 сетки df2ed4841a9453ca
// Назначение: тест Matrix_PSLL101Override_DemandBackRestartsConfirm набора FB_CemGen01_Test
//             (сценарий по матрице, DESIGN.md, 12.4).
// Автор:      kr0nsch; код — генератор cemgen
// Версия:     1.0.0
// Документ:   docs/DESIGN.md, раздел «10. Генератор cemgen»; docs/cause_effect_matrix.md
// ВНИМАНИЕ:   код демонстрационный и не предназначен для систем безопасности. Реальная ПАЗ требует
//             определения SIL, сертифицированных аппаратных и программных средств и валидации по
//             ГОСТ Р МЭК 61511.
// Причина 2 PSLL101: пусковой обход и требование в t0; норма с t1; ровно на t1 + 30 с, когда обход
// снялся бы, требование снова — обход действует, подтверждение нормы сброшено; норма с t2; на t2 + 30
// с − шаг обход действует; на t2 + 30 с — OverrideCleared.
METHOD PRIVATE PSLL101OverrideDemandBackRestartsConfirm
VAR
    xArmed : BOOL;   // стенд взведён: все следствия под напряжением после сброса
END_VAR

(* ---- PSLL101OverrideExpiresThenTrips.method.decl.st ---- *)
// AUTO-GENERATED by cemgen 1.0.0 — не редактировать: правьте матрицу и запустите
//   python -m cemgen generate <файл матрицы .csv или .xlsx>
// Матрица: SIS-V101-CEM, объект V-101, ревизия B от 2026-10-19, SHA-256 сетки df2ed4841a9453ca
// Назначение: тест Matrix_PSLL101Override_ExpiresThenTrips набора FB_CemGen01_Test (сценарий по
//             матрице, DESIGN.md, 12.4).
// Автор:      kr0nsch; код — генератор cemgen
// Версия:     1.0.0
// Документ:   docs/DESIGN.md, раздел «10. Генератор cemgen»; docs/cause_effect_matrix.md
// ВНИМАНИЕ:   код демонстрационный и не предназначен для систем безопасности. Реальная ПАЗ требует
//             определения SIL, сертифицированных аппаратных и программных средств и валидации по
//             ГОСТ Р МЭК 61511.
// Причина 2 PSLL101: ключ разрешения обходов, запрос пускового обхода и требование в одном вызове t0;
// до t0 + 15 мин − шаг обход действует, причина не зафиксирована; ровно на t0 + 15 мин —
// OverrideExpired, фиксация, первопричина PSLL101.
METHOD PRIVATE PSLL101OverrideExpiresThenTrips
VAR
    xArmed : BOOL;   // стенд взведён: все следствия под напряжением после сброса
END_VAR

(* ---- PSLL101OverrideExpiryBoundsConfirm.method.decl.st ---- *)
// AUTO-GENERATED by cemgen 1.0.0 — не редактировать: правьте матрицу и запустите
//   python -m cemgen generate <файл матрицы .csv или .xlsx>
// Матрица: SIS-V101-CEM, объект V-101, ревизия B от 2026-10-19, SHA-256 сетки df2ed4841a9453ca
// Назначение: тест Matrix_PSLL101Override_ExpiryBoundsConfirm набора FB_CemGen01_Test (сценарий по
//             матрице, DESIGN.md, 12.4).
// Автор:      kr0nsch; код — генератор cemgen
// Версия:     1.0.0
// Документ:   docs/DESIGN.md, раздел «10. Генератор cemgen»; docs/cause_effect_matrix.md
// ВНИМАНИЕ:   код демонстрационный и не предназначен для систем безопасности. Реальная ПАЗ требует
//             определения SIL, сертифицированных аппаратных и программных средств и валидации по
//             ГОСТ Р МЭК 61511.
// Причина 2 PSLL101: пусковой обход и требование в t0; норма с t0 + 14 мин 30 с + шаг — подтверждение
// (30 с) закончилось бы после срока; на t0 + 15 мин − шаг обход действует; ровно на t0 + 15 мин —
// OverrideExpired (срок — верхняя граница), OverrideCleared нет, причина не зафиксирована (требования
// нет).
METHOD PRIVATE PSLL101OverrideExpiryBoundsConfirm
VAR
    xArmed : BOOL;   // стенд взведён: все следствия под напряжением после сброса
END_VAR

(* ---- PSLL101ResetOnlyAfterClear.method.decl.st ---- *)
// AUTO-GENERATED by cemgen 1.0.0 — не редактировать: правьте матрицу и запустите
//   python -m cemgen generate <файл матрицы .csv или .xlsx>
// Матрица: SIS-V101-CEM, объект V-101, ревизия B от 2026-10-19, SHA-256 сетки df2ed4841a9453ca
// Назначение: тест Matrix_PSLL101Reset_OnlyAfterClear набора FB_CemGen01_Test (сценарий по матрице,
//             DESIGN.md, 12.4).
// Автор:      kr0nsch; код — генератор cemgen
// Версия:     1.0.0
// Документ:   docs/DESIGN.md, раздел «10. Генератор cemgen»; docs/cause_effect_matrix.md
// ВНИМАНИЕ:   код демонстрационный и не предназначен для систем безопасности. Реальная ПАЗ требует
//             определения SIL, сертифицированных аппаратных и программных средств и валидации по
//             ГОСТ Р МЭК 61511.
// Причина 2 PSLL101: срабатывание; сброс при требовании → ResetDenied, блокирует PSLL101, следствия
// обесточены; норма → следствия всё ещё обесточены (фиксация); сброс → все следствия под напряжением.
METHOD PRIVATE PSLL101ResetOnlyAfterClear
VAR
    xArmed : BOOL;          // стенд взведён: все следствия под напряжением после сброса
    stEv   : ST_SisEvent;   // последнее событие журнала
END_VAR

(* ---- TSHH103BypassExpiresBackToVoting.method.decl.st ---- *)
// AUTO-GENERATED by cemgen 1.0.0 — не редактировать: правьте матрицу и запустите
//   python -m cemgen generate <файл матрицы .csv или .xlsx>
// Матрица: SIS-V101-CEM, объект V-101, ревизия B от 2026-10-19, SHA-256 сетки df2ed4841a9453ca
// Назначение: тест Matrix_TSHH103Bypass_ExpiresBackToVoting набора FB_CemGen01_Test (сценарий по
//             матрице, DESIGN.md, 12.4).
// Автор:      kr0nsch; код — генератор cemgen
// Версия:     1.0.0
// Документ:   docs/DESIGN.md, раздел «10. Генератор cemgen»; docs/cause_effect_matrix.md
// ВНИМАНИЕ:   код демонстрационный и не предназначен для систем безопасности. Реальная ПАЗ требует
//             определения SIL, сертифицированных аппаратных и программных средств и валидации по
//             ГОСТ Р МЭК 61511.
// Причина 5 TSHH103: ключ разрешения байпасов, байпас TT103A → Active; канал недостоверен → Bypassed,
// не сработало; на t0 + 8 ч − шаг — Active; ровно на t0 + 8 ч — Expired, BypassExpired, канал Invalid;
// далее — по эталонной модели.
METHOD PRIVATE TSHH103BypassExpiresBackToVoting
VAR
    xArmed : BOOL;           // стенд взведён: все следствия под напряжением после сброса
    stVs   : ST_VotingSts;   // копия состояния группы голосования
END_VAR

(* ---- TSHH103ChannelInvalidMatchesPolicy.method.decl.st ---- *)
// AUTO-GENERATED by cemgen 1.0.0 — не редактировать: правьте матрицу и запустите
//   python -m cemgen generate <файл матрицы .csv или .xlsx>
// Матрица: SIS-V101-CEM, объект V-101, ревизия B от 2026-10-19, SHA-256 сетки df2ed4841a9453ca
// Назначение: тест Matrix_TSHH103ChannelInvalid_MatchesPolicy набора FB_CemGen01_Test (сценарий по
//             матрице, DESIGN.md, 12.4).
// Автор:      kr0nsch; код — генератор cemgen
// Версия:     1.0.0
// Документ:   docs/DESIGN.md, раздел «10. Генератор cemgen»; docs/cause_effect_matrix.md
// ВНИМАНИЕ:   код демонстрационный и не предназначен для систем безопасности. Реальная ПАЗ требует
//             определения SIL, сертифицированных аппаратных и программных средств и валидации по
//             ГОСТ Р МЭК 61511.
// Причина 5 TSHH103 (1oo2, DegradeSafe): канал TT103A недостоверен → действующая схема и срабатывание
// по политике деградации; если не сработало — требование на TT103B → по эталонной модели.
METHOD PRIVATE TSHH103ChannelInvalidMatchesPolicy
VAR
    xArmed : BOOL;           // стенд взведён: все следствия под напряжением после сброса
    stVs   : ST_VotingSts;   // копия состояния группы голосования
END_VAR

(* ---- TSHH103DelayTripsExactlyAtDelay.method.decl.st ---- *)
// AUTO-GENERATED by cemgen 1.0.0 — не редактировать: правьте матрицу и запустите
//   python -m cemgen generate <файл матрицы .csv или .xlsx>
// Матрица: SIS-V101-CEM, объект V-101, ревизия B от 2026-10-19, SHA-256 сетки df2ed4841a9453ca
// Назначение: тест Matrix_TSHH103Delay_TripsExactlyAtDelay набора FB_CemGen01_Test (сценарий по
//             матрице, DESIGN.md, 12.4).
// Автор:      kr0nsch; код — генератор cemgen
// Версия:     1.0.0
// Документ:   docs/DESIGN.md, раздел «10. Генератор cemgen»; docs/cause_effect_matrix.md
// ВНИМАНИЕ:   код демонстрационный и не предназначен для систем безопасности. Реальная ПАЗ требует
//             определения SIL, сертифицированных аппаратных и программных средств и валидации по
//             ГОСТ Р МЭК 61511.
// Причина 5 TSHH103: требование в t0; на t0 + 5 с − шаг не зафиксирована, следствия под напряжением;
// ровно на t0 + 5 с — зафиксирована, ltFirstOut = t0 + задержка.
METHOD PRIVATE TSHH103DelayTripsExactlyAtDelay
VAR
    xArmed : BOOL;    // стенд взведён: все следствия под напряжением после сброса
    ltT0   : LTIME;   // момент t0 по подменному времени стенда
END_VAR

(* ---- TSHH103DemandTripsOwnEffects.method.decl.st ---- *)
// AUTO-GENERATED by cemgen 1.0.0 — не редактировать: правьте матрицу и запустите
//   python -m cemgen generate <файл матрицы .csv или .xlsx>
// Матрица: SIS-V101-CEM, объект V-101, ревизия B от 2026-10-19, SHA-256 сетки df2ed4841a9453ca
// Назначение: тест Matrix_TSHH103Demand_TripsOwnEffects набора FB_CemGen01_Test (сценарий по
//             матрице, DESIGN.md, 12.4).
// Автор:      kr0nsch; код — генератор cemgen
// Версия:     1.0.0
// Документ:   docs/DESIGN.md, раздел «10. Генератор cemgen»; docs/cause_effect_matrix.md
// ВНИМАНИЕ:   код демонстрационный и не предназначен для систем безопасности. Реальная ПАЗ требует
//             определения SIL, сертифицированных аппаратных и программных средств и валидации по
//             ГОСТ Р МЭК 61511.
// Причина 5 TSHH103 (1oo2, задержка 5 с): требование TT103A, TT103B = 13,23 мА (86,5 °C; уставка ≥ 85
// °C) отключает H101, UA110; остальные следствия под напряжением; первопричина TSHH103.
METHOD PRIVATE TSHH103DemandTripsOwnEffects
VAR
    xArmed : BOOL;   // стенд взведён: все следствия под напряжением после сброса
END_VAR

(* ---- TSHH103OverrideDenied.method.decl.st ---- *)
// AUTO-GENERATED by cemgen 1.0.0 — не редактировать: правьте матрицу и запустите
//   python -m cemgen generate <файл матрицы .csv или .xlsx>
// Матрица: SIS-V101-CEM, объект V-101, ревизия B от 2026-10-19, SHA-256 сетки df2ed4841a9453ca
// Назначение: тест Matrix_TSHH103Override_Denied набора FB_CemGen01_Test (сценарий по матрице,
//             DESIGN.md, 12.4).
// Автор:      kr0nsch; код — генератор cemgen
// Версия:     1.0.0
// Документ:   docs/DESIGN.md, раздел «10. Генератор cemgen»; docs/cause_effect_matrix.md
// ВНИМАНИЕ:   код демонстрационный и не предназначен для систем безопасности. Реальная ПАЗ требует
//             определения SIL, сертифицированных аппаратных и программных средств и валидации по
//             ГОСТ Р МЭК 61511.
// Причина 5 TSHH103 без разрешённого обхода: ключ разрешения обходов, запрос → последнее событие
// OverrideDenied, обхода нет; требование → срабатывание после задержки.
METHOD PRIVATE TSHH103OverrideDenied
VAR
    xArmed : BOOL;          // стенд взведён: все следствия под напряжением после сброса
    stEv   : ST_SisEvent;   // последнее событие журнала
END_VAR

(* ---- TSHH103ResetOnlyAfterClear.method.decl.st ---- *)
// AUTO-GENERATED by cemgen 1.0.0 — не редактировать: правьте матрицу и запустите
//   python -m cemgen generate <файл матрицы .csv или .xlsx>
// Матрица: SIS-V101-CEM, объект V-101, ревизия B от 2026-10-19, SHA-256 сетки df2ed4841a9453ca
// Назначение: тест Matrix_TSHH103Reset_OnlyAfterClear набора FB_CemGen01_Test (сценарий по матрице,
//             DESIGN.md, 12.4).
// Автор:      kr0nsch; код — генератор cemgen
// Версия:     1.0.0
// Документ:   docs/DESIGN.md, раздел «10. Генератор cemgen»; docs/cause_effect_matrix.md
// ВНИМАНИЕ:   код демонстрационный и не предназначен для систем безопасности. Реальная ПАЗ требует
//             определения SIL, сертифицированных аппаратных и программных средств и валидации по
//             ГОСТ Р МЭК 61511.
// Причина 5 TSHH103: срабатывание; сброс при требовании → ResetDenied, блокирует TSHH103, следствия
// обесточены; норма → следствия всё ещё обесточены (фиксация); сброс → все следствия под напряжением.
METHOD PRIVATE TSHH103ResetOnlyAfterClear
VAR
    xArmed : BOOL;          // стенд взведён: все следствия под напряжением после сброса
    stEv   : ST_SisEvent;   // последнее событие журнала
END_VAR
